TYPE ST_PolarIIChamber_ArmAlignTestParam :
STRUCT
	ArmIndex : UINT; // 1..4
	NozzleIndex : UINT; // 1..3
	Recipe : ST_PolarIIChamber_Recipe;
	TestTime : TIME;
END_STRUCT
END_TYPE

(* stored: Version 1.1.0.1, ProductVersion 3.1.4026.18
   DUT ST_PolarIIChamber_ArmAlignTestParam: Id {14000000-0000-0000-0000-000000000016} *)
